(* IEC 61131-3 sources: kns-port-domestic/upstream/kns-pump-station/src/POUs/Station/FB_LevelControlStepped, 2 files *)

(* ---- FB_LevelControlStepped.decl.st ---- *)
// Назначение: ступенчатое регулирование по уровням пуска и останова с гистерезисом (04 §6):
//             автомат 0/1/2 насоса, каждое пересечение подтверждается выдержкой tLvlConfirm
//             (границы включительно: пуск при уровне >=, останов при <=). Недостоверный уровень —
//             состояние держится. При xEnable = FALSE выход 0, автомат работает дальше (таймеры
//             непрерывны), состояние задаёт следующий xInit (вход без рывка по числу работающих).
// Автор:      kr0nsch
// Версия:     0.1.0
// Документ:   docs/DESIGN.md, раздел 6.3; docs/04_algorithms.md, раздел 6
FUNCTION_BLOCK FB_LevelControlStepped
VAR_INPUT
    xEnable     : BOOL;             // eControlAct = Stepped
    rLevel_m    : REAL;             // fbLT101.rValue_eu
    xLevelValid : BOOL;             // fbLT101.xValid
    xInit       : BOOL;             // импульс: число насосов := uiInitPumps (вход без рывка)
    uiInitPumps : UINT;             // работающие насосы станции
    itfTime     : PL.I_TimeSource;
END_VAR
VAR_IN_OUT CONSTANT
    stCfg : ST_StationCfg;          // rLvl*_m, tLvlConfirm, rStepSpeed_pct, uiDutyMax
END_VAR
VAR_OUTPUT
    uiRequired  : UINT;             // 0…MIN(2, uiDutyMax)
    rSpeed_pct  : REAL;             // stCfg.rStepSpeed_pct
    xConfirming : BOOL;             // идёт выдержка tLvlConfirm
END_VAR
VAR
    uiPumps        : UINT;          // состояние автомата: 0, 1, 2 насоса
    fbStartLead    : PL.FB_Delay;   // 0 → 1: уровень >= rLvlStartLead_m
    fbStartAssist  : PL.FB_Delay;   // 1 → 2: уровень >= rLvlStartAssist_m
    fbStopAssist   : PL.FB_Delay;   // 2 → 1: уровень <= rLvlStopAssist_m
    fbStopAll      : PL.FB_Delay;   // 1, 2 → 0: уровень <= rLvlStop_m
END_VAR
VAR_TEMP
    uiMax : UINT;                   // предел числа насосов: MIN(STN_DUTY_MAX, uiDutyMax)
END_VAR

(* ---- FB_LevelControlStepped.impl.st ---- *)
// Ступенчатый способ — не больше двух насосов (ведущий и подпорный) и не больше uiDutyMax
uiMax := MIN(GVL_Const.STN_DUTY_MAX, stCfg.uiDutyMax);

// 1. Вход без рывка: число насосов — по работающим; выдержки подтверждения — заново
IF xInit THEN
    uiPumps := MIN(uiInitPumps, uiMax);
    fbStartLead.Preset(xValue := FALSE);
    fbStartAssist.Preset(xValue := FALSE);
    fbStopAssist.Preset(xValue := FALSE);
    fbStopAll.Preset(xValue := FALSE);
END_IF
uiPumps := MIN(uiPumps, uiMax);

// 2. Пересечения уровней по диаграмме 04 §6. Условие каждого перехода зависит от состояния: после
//    перехода выдержка следующего начинается заново. Недостоверный уровень — условий нет, состояние
//    держится (сравнения с NaN ложны и без проверки xLevelValid)
fbStartLead(xIn := xLevelValid AND uiPumps = 0 AND rLevel_m >= stCfg.rLvlStartLead_m AND uiMax > 0,
            tOnDelay := stCfg.tLvlConfirm, itfTime := itfTime);
fbStartAssist(xIn := xLevelValid AND uiPumps = 1 AND rLevel_m >= stCfg.rLvlStartAssist_m AND uiMax > 1,
              tOnDelay := stCfg.tLvlConfirm, itfTime := itfTime);
fbStopAssist(xIn := xLevelValid AND uiPumps = 2 AND rLevel_m <= stCfg.rLvlStopAssist_m,
             tOnDelay := stCfg.tLvlConfirm, itfTime := itfTime);
fbStopAll(xIn := xLevelValid AND uiPumps > 0 AND rLevel_m <= stCfg.rLvlStop_m,
          tOnDelay := stCfg.tLvlConfirm, itfTime := itfTime);

// 3. Переход: останов всех старше остальных (2 → 0 одним шагом, если обе выдержки истекли)
IF fbStopAll.xOut THEN
    uiPumps := 0;
ELSIF fbStopAssist.xOut THEN
    uiPumps := 1;
ELSIF fbStartAssist.xOut THEN
    uiPumps := 2;
ELSIF fbStartLead.xOut THEN
    uiPumps := 1;
END_IF

xConfirming := fbStartLead.xTimingOn OR fbStartAssist.xTimingOn OR fbStopAssist.xTimingOn
               OR fbStopAll.xTimingOn;
uiRequired := SEL(xEnable, 0, uiPumps);
rSpeed_pct := stCfg.rStepSpeed_pct;
